FUNCTION_BLOCK FB_SystemSM
VAR_INPUT
END_VAR
VAR_OUTPUT
END_VAR
VAR
END_VAR

// Edge-Detect Commands
// MOVE ME!!
//_TrigStart(CLK := HMI.bStart);
//_TrigStop(CLK := HMI.bStop);
//_TrigReset(CLK := HMI.bReset);

END_FUNCTION_BLOCK

(* stored: Version 1.1.0.1
   POU FB_SystemSM: Id {41c29ac7-c7f9-4bcc-9f26-f0832b5cf229}, SpecialFunc None *)
